// TIA Portal V21 export
// export: Created 2026-10-23T20:42:14.793557Z, ExportSetting WithDefaults, DisplayName Totally Integrated Automation Portal, DisplayVersion V21 Update 1, DisplayName SINAMICS Startdrive Advanced, DisplayVersion V21 HF2, DisplayName SINAMICS Startdrive G110M, G120, G120C, G120D, G120P, G115D, DisplayVersion V21 HF2, DisplayName SINAMICS Startdrive G130, G150, S120, S150, G200, G220, S200, S210, S220, Innomotics MVD, DisplayVersion V21 HF2, DisplayName STEP 7 Professional, DisplayVersion V21 Update 1, DisplayName STEP 7 Safety, DisplayVersion V21, DisplayName Tech WebApplication, DisplayVersion V21, DisplayName WinCC Basic/Comfort/Advanced, DisplayVersion V21 Update 1, DisplayName WinCC Unified, DisplayVersion V21 Update 1
FUNCTION "F_FC_Logic" : Void   // FC9, F_FBD
{ S7_Optimized_Access := 'TRUE' }
VERSION : 0.1
// stored: AutoNumber true, IsIECCheckEnabled false, UDAEnableTagReadback false
   VAR_INPUT
      GuardClosed : Bool;   // Schutztür geschlossen / Guard door closed
      SetupMode : Bool;   // Einrichtbetrieb angewählt / Setup mode selected
      EmergencyStopOk : Bool;   // Not-Halt nicht betätigt / Emergency stop not pressed
   END_VAR
   VAR_OUTPUT
      Release : Bool;   // Freigabe der Maschine / Release of the machine
   END_VAR
BEGIN

REGION Network 1: Schutztür oder Einrichtbetrieb, und Not-Halt in Ordnung / Guard or setup mode, and emergency stop ok
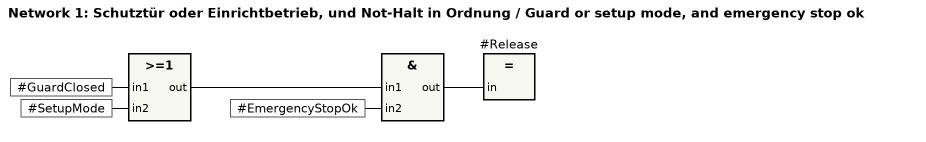
   #Release := (#GuardClosed OR #SetupMode) AND #EmergencyStopOk;
END_REGION
END_FUNCTION
